// TIA Portal V20 export
Screen "Pop-up_ISRA VISION"  395x450
  ScreenItem "Robot Name" at 2,2 size 393x48  Type=HmiIOField
  ScreenItem "Background" at -1,49 size 395x400  Type=HmiRectangle
  ScreenItem "Cancel Mode" at 315,4 size 76x42  Type=HmiButton
  ScreenItem "矩形_4" at 29,85 size 324x354  Type=HmiRectangle
  ScreenItem "Text Field In Auto On_9" at 41,121 size 148x21  Type=HmiTextBox
  ScreenItem "Text Field Home Position_17" at 41,145 size 148x21  Type=HmiTextBox
  ScreenItem "Text field Robot Status_5" at 31,86 size 324x30  Type=HmiTextBox
  ScreenItem "Text Field System Ready_9" at 41,169 size 148x21  Type=HmiTextBox
  ScreenItem "Text Field Motor On_9" at 41,193 size 148x21  Type=HmiTextBox
  ScreenItem "Text Field Home Position_18" at 196,121 size 148x21  Type=HmiTextBox
  ScreenItem "Text Field Manual_18" at 196,193 size 148x21  Type=HmiTextBox
  ScreenItem "Text Field Cycle On_18" at 196,145 size 148x21  Type=HmiTextBox
  ScreenItem "Text Field On Path_18" at 196,169 size 148x21  Type=HmiTextBox
  ScreenItem "FaultNo" at 189,249 size 108x63  Type=HmiIOField
  ScreenItem "Text field_8" at 87,266 size 94x29  Type=HmiTextBox
